(* Logix 5000 project; controller DSFW_Budzar vendor 1 type 14 code 154 rev 32.13; software revision 32.03; part 3 of 5 *)
(* tags used below, declared in another part *)
   ALARMS : DINT[5];
   ALWAYS_OFF : BOOL;
   Batch_Mode_Enable : BOOL;
   BudLib_P2T_1 : BudLib_Superheat_Subcooling;
   BudLib_P2T_2 : BudLib_Superheat_Subcooling;
   BudLib_P2T_3 : BudLib_Superheat_Subcooling;
   CLR_Alarms : BOOL;
   Compressor_R404A_Subcooling : REAL;
   Compressor_R404A_Superheat : REAL;
   CR_108 : ALIAS FOR Local:1:O.Data.0;   // Process Pump Motor Relay (Energizes Contactor M-101)
   CR_109 : ALIAS FOR Local:1:O.Data.5;   // Compressor Motor Relay (Energizes Contactor C-101)
   CR_201 : ALIAS FOR Local:1:O.Data.8;   // GFS-10 Auto Start Relay (Enables Glycol Pump)
   Enable_Batch : BOOL;   // Batch/Jacket Mode 0=Jacket 1=Batch
   Evaporator_R404A_Superheat : REAL;
   F8 : REAL[48];   // FLOAT DATA FOR PLANT SUPERVISORY SYSTEM
   FIC_101_Run_PID : BOOL;
   FIC_101_Stop_PID : BOOL;
   FIT_101 : BL_Analog_Input;   // Flow Indicating Transmitter
   FIT_101_PID_Scale_Max : REAL;
   FIT_101_PID_Scale_Min : REAL;
   Glycol_Pump_Disable_TMR : TIMER;   // Disable Glycol Fill Pump on High PSI (backup for Pressure Switch on Neptune)
   HMI_Bypass_Speed : DINT;
   HMI_Bypass_Status : BOOL;
   HMI_FCV_101_CV : REAL;
   HMI_Heater_1_Lamp : BOOL;
   HMI_Pump_Start : BOOL;
   HMI_Pump_Status : BOOL;
   HMI_Pump_Stop : BOOL;
   HMI_Ramping : BOOL;
   HMI_SCR_Max : DINT;
   HMI_Soaking : BOOL;
   HMI_Supply_Flow_Speed : DINT;
   HMI_Supply_Flow_Status : BOOL;
   Local_System_Start : BOOL;   // Local System Start 0=Stop 1=Start
   Local_Temp_Setpoint : REAL;   // Local Temperature Setpoint
   M_101_AUX : ALIAS FOR Local:1:I.Data.3;
   ONS : DINT[3];   // One-Shots
   PLC_DateTime : DINT[7];
   PM_101 : ALIAS FOR Local:1:I.Data.1;
   PT_101 : BL_Analog_Input;   // Process Supply Pressure
   PT_102 : BL_Analog_Input;   // R404A Compressor Suction Pressure
   PT_102_PID_Scale_Max : REAL;
   PT_102_PID_Scale_Min : REAL;
   PT_103 : BL_Analog_Input;   // R404A Compressor Discharge Pressure
   PT_103_PID_Scale_Max : REAL;
   PT_103_PID_Scale_Min : REAL;
   PT_104 : BL_Analog_Input;   // R404A Evaporator Suction Pressure
   PT_104_PID_Scale_Max : REAL;
   PT_104_PID_Scale_Min : REAL;
   PT_105 : BL_Analog_Input;   // Condenser Chilled Glycol Return Pressure
   PT_106 : BL_Analog_Input;   // Condenser Chilled Glycol Supply Pressure
   PT_107 : BL_Analog_Input;   // Process Pump Suction Pressure
   PT_108 : BL_Analog_Input;   // Process Pump Suction Discharge Pressure
   Pump_Manual_Release : BOOL;
   Pump_Manual_Release_Timer : TIMER;
   Pump_OK_To_Run : BOOL;
   REACTOR_BATCH_PID_START : BOOL;
   REACTOR_BATCH_PID_STOP : BOOL;
   REACTOR_BATCH_PIDE : PID_ENHANCED;
   REACTOR_BATCH_PV : REAL;
   REACTOR_BATCH_SP_HIGH : REAL;
   REACTOR_BATCH_SP_LOW : REAL;
   REACTOR_HEAT_RUN_PIDE : BOOL;
   REACTOR_HEAT_STOP_PIDE : BOOL;
   REACTOR_HEATERS_OK_TO_RUN : BOOL;
   REACTOR_HEATERS_TEMPERATURE_PIDE : PID_ENHANCED;
   Remote_Enable_Batch : BOOL;   // Remote Jacket/Batch Control (0=Jacket, 1=Batch)
   Remote_System_Start : BOOL;   // Remote Start/Stop 0=Stop 1=Start
   Remote_Temp_Setpoint : REAL;   // Remote Temperature Setpoint
   RX_Profile_Stop_SP_Control : TIMER;
   RX_RMPS : RAMP_SOAK;
   RX_RMPS_Current_Segment : DINT;
   RX_RMPS_Output : REAL;
   RX_RMPS_Soak_Time : REAL[11];
   RX_RMPS_Soak_Value : REAL[11];
   RX_RMPS_SP_Out : REAL;
   RX_Run_Temp_Profile : BOOL;
   RX_Start_Temperature_Profile : BOOL;
   RX_Stop_Temp_Profile : BOOL;
   SCR_Output_Percent : DINT;
   SCR_PID_Request : REAL;
   Sensor_1 : BudLib_Analog_Sensor;
   Sensor_2 : BudLib_Analog_Sensor;
   Sensor_3 : BudLib_Analog_Sensor;
   Sensor_4 : BudLib_Analog_Sensor;
   Sensor_5 : BudLib_Analog_Sensor;
   Sensor_6 : BudLib_Analog_Sensor;
   Sensor_7 : BudLib_Analog_Sensor;
   Sensor_8 : BudLib_Analog_Sensor;
   Sensor_9 : BudLib_Analog_Sensor;
   System_Mode : BOOL;   // 0 = Local Control 1 = Remote Control
   System_Start : BOOL;   // System Start
   T_SENSOR_1 : BudLib_Analog_Sensor;
   T_SENSOR_2 : BudLib_Analog_Sensor;
   T_SENSOR_3 : BudLib_Analog_Sensor;
   T_SENSOR_4 : BudLib_Analog_Sensor;
   T_SENSOR_5 : BudLib_Analog_Sensor;
   T_SENSOR_6 : BudLib_Analog_Sensor;
   T_SENSOR_8 : BudLib_Analog_Sensor;
   TE_101 : BL_Analog_Input;   // Process Supply Temperature
   TE_102 : BL_Analog_Input;   // Process Return Temperature
   TE_103 : BL_Analog_Input;   // R507A Liquid Line Temperature
   TE_104 : BL_Analog_Input;   // R507A Evaporator Suction Temperature
   TE_105 : BL_Analog_Input;   // R507A Compressor Suction Temperature
   TE_106 : BL_Analog_Input;   // CONDENSER CHILLED GLYCOL OUTLET TEMPERATURE SENSOR
   TE_108 : BL_Analog_Input;   // CONDENSER CHILLED GLYCOL INLET TEMPERATURE SENSOR
   Temperature_Setpoint : REAL;
   Temperature_Setpoint_Max : REAL;   // Maximum Operating Temperature Setpoint (Deg C)
   Temperature_Setpoint_Min : REAL;   // Minimum Operating Temperature Setpoint (Deg C)
   TSH_101 : ALIAS FOR Local:1:I.Data.4;
   VESSEL_TEMPERATURE : BL_Analog_Input;   // End User Reactor Temperature
(* A_MainProgram, continued *)

ROUTINE Routine_Schedule   (* ladder *)
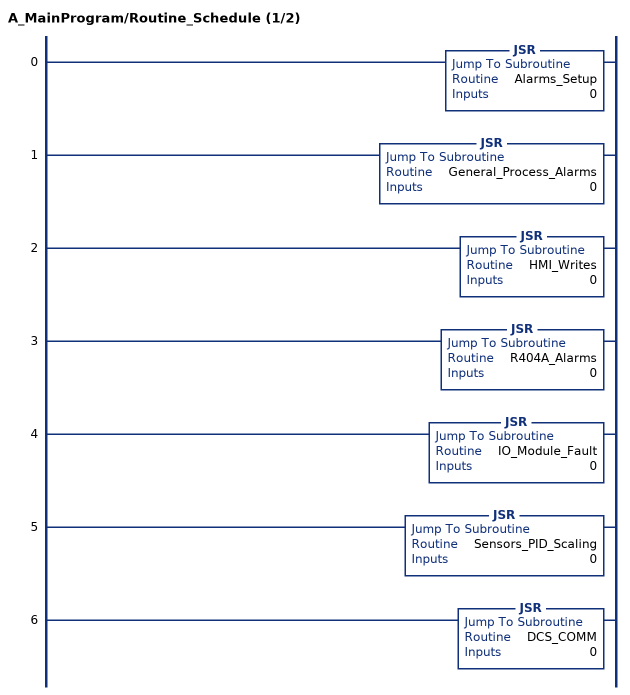
   0: JSR(Alarms_Setup,0);
   1: JSR(General_Process_Alarms,0);
   2: JSR(HMI_Writes,0);
   3: JSR(R404A_Alarms,0);
   4: JSR(IO_Module_Fault,0);
   5: JSR(Sensors_PID_Scaling,0);
   6: JSR(DCS_COMM,0);
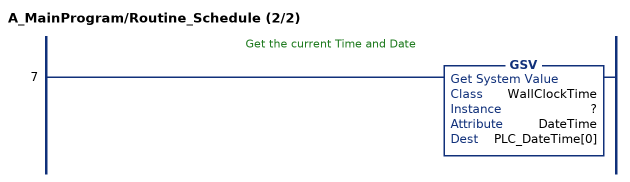
   // Get the current Time and Date
   7: GSV(WallClockTime,?,DateTime,PLC_DateTime[0]);
END_ROUTINE

ROUTINE Sensors_PID_Scaling   (* ladder *)
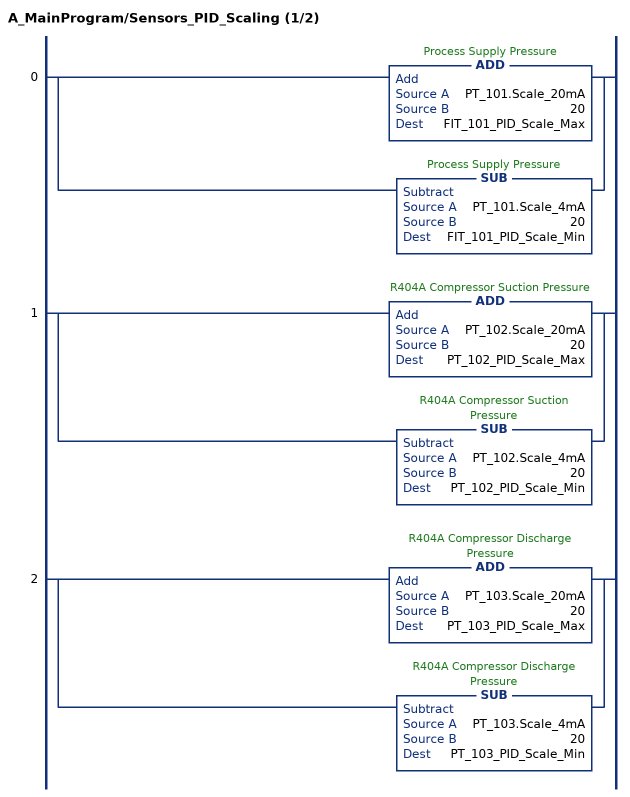
   0: [ADD(PT_101.Scale_20mA,20,FIT_101_PID_Scale_Max) ,SUB(PT_101.Scale_4mA,20,FIT_101_PID_Scale_Min) ];
   1: [ADD(PT_102.Scale_20mA,20,PT_102_PID_Scale_Max) ,SUB(PT_102.Scale_4mA,20,PT_102_PID_Scale_Min) ];
   2: [ADD(PT_103.Scale_20mA,20,PT_103_PID_Scale_Max) ,SUB(PT_103.Scale_4mA,20,PT_103_PID_Scale_Min) ];
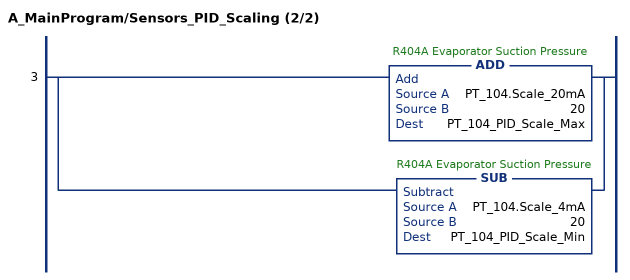
   3: [ADD(PT_104.Scale_20mA,20,PT_104_PID_Scale_Max) ,SUB(PT_104.Scale_4mA,20,PT_104_PID_Scale_Min) ];
END_ROUTINE
END_PROGRAM

PROGRAM B_Process_Control   (* main routine Main *)
VAR
   test_th : BOOL;
END_VAR

ROUTINE A_Sensors   (* ladder *)
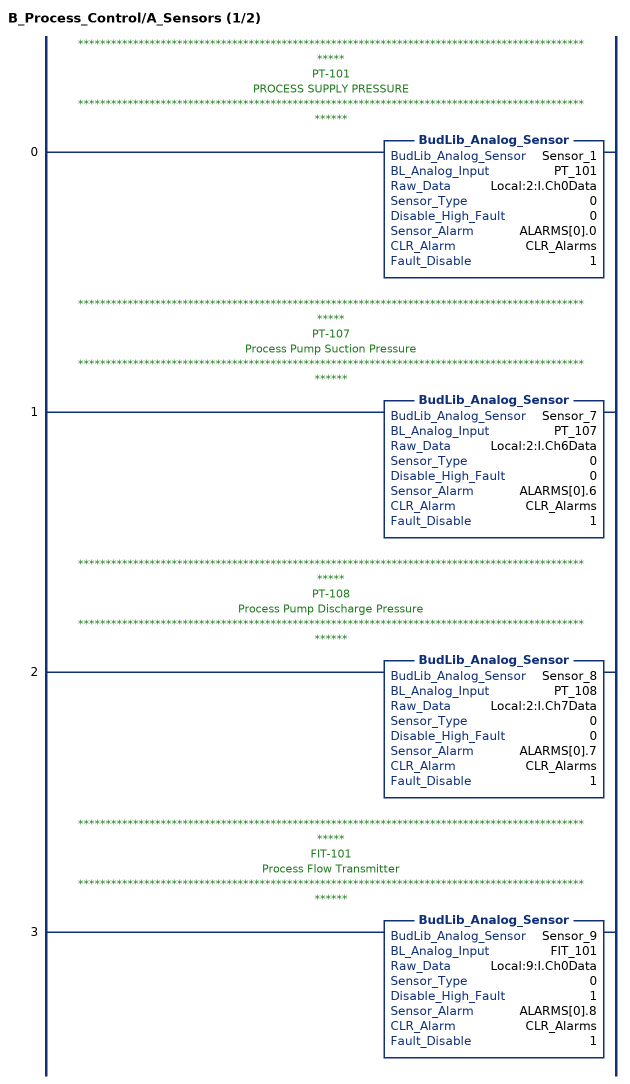
   // *************************************************************************************************
   // PT-101
   // PROCESS SUPPLY PRESSURE
   // **************************************************************************************************
   0: BudLib_Analog_Sensor(Sensor_1,PT_101,Local:2:I.Ch0Data,0,0,ALARMS[0].0,CLR_Alarms,1);
   // *************************************************************************************************
   // PT-107
   // Process Pump Suction Pressure
   // **************************************************************************************************
   1: BudLib_Analog_Sensor(Sensor_7,PT_107,Local:2:I.Ch6Data,0,0,ALARMS[0].6,CLR_Alarms,1);
   // *************************************************************************************************
   // PT-108
   // Process Pump Discharge Pressure
   // **************************************************************************************************
   2: BudLib_Analog_Sensor(Sensor_8,PT_108,Local:2:I.Ch7Data,0,0,ALARMS[0].7,CLR_Alarms,1);
   // *************************************************************************************************
   // FIT-101
   // Process Flow Transmitter
   // **************************************************************************************************
   3: BudLib_Analog_Sensor(Sensor_9,FIT_101,Local:9:I.Ch0Data,0,1,ALARMS[0].8,CLR_Alarms,1);
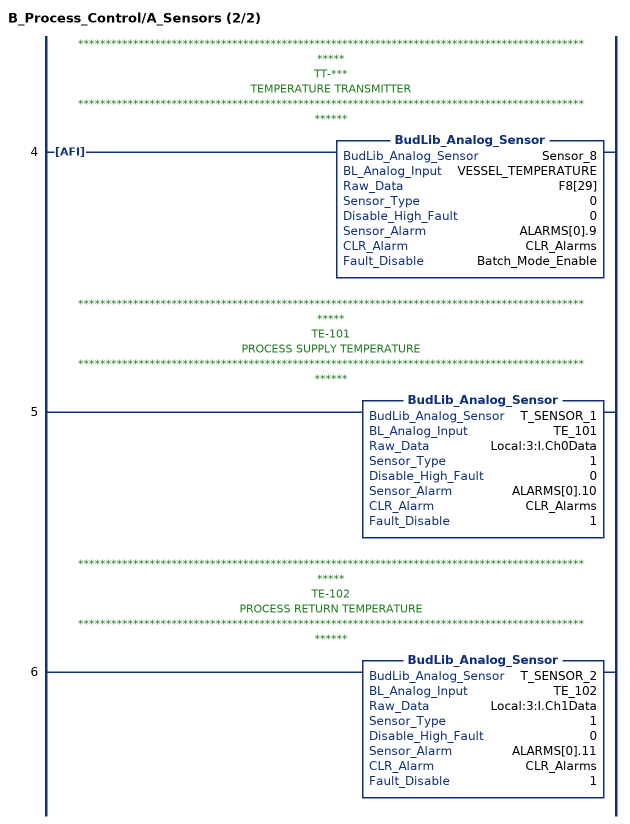
   // *************************************************************************************************
   // TT-***
   // TEMPERATURE TRANSMITTER
   // **************************************************************************************************
   4: AFI()BudLib_Analog_Sensor(Sensor_8,VESSEL_TEMPERATURE,F8[29],0,0,ALARMS[0].9,CLR_Alarms,Batch_Mode_Enable);
   // *************************************************************************************************
   // TE-101
   // PROCESS SUPPLY TEMPERATURE
   // **************************************************************************************************
   5: BudLib_Analog_Sensor(T_SENSOR_1,TE_101,Local:3:I.Ch0Data,1,0,ALARMS[0].10,CLR_Alarms,1);
   // *************************************************************************************************
   // TE-102
   // PROCESS RETURN TEMPERATURE
   // **************************************************************************************************
   6: BudLib_Analog_Sensor(T_SENSOR_2,TE_102,Local:3:I.Ch1Data,1,0,ALARMS[0].11,CLR_Alarms,1);
END_ROUTINE

ROUTINE Glycol_Tank   (* ladder *)
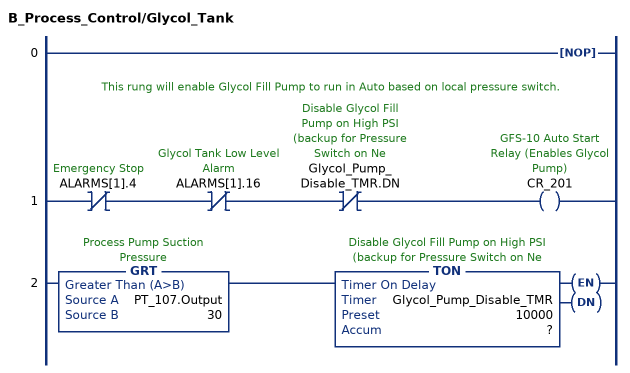
   0: NOP();
   // This rung will enable Glycol Fill Pump to run in Auto based on local pressure switch.
   1: XIO(ALARMS[1].4)XIO(ALARMS[1].16)XIO(Glycol_Pump_Disable_TMR.DN)OTE(CR_201);
   2: GRT(PT_107.Output,30)TON(Glycol_Pump_Disable_TMR,?,?);
END_ROUTINE

ROUTINE Heaters_Control   (* ladder *)
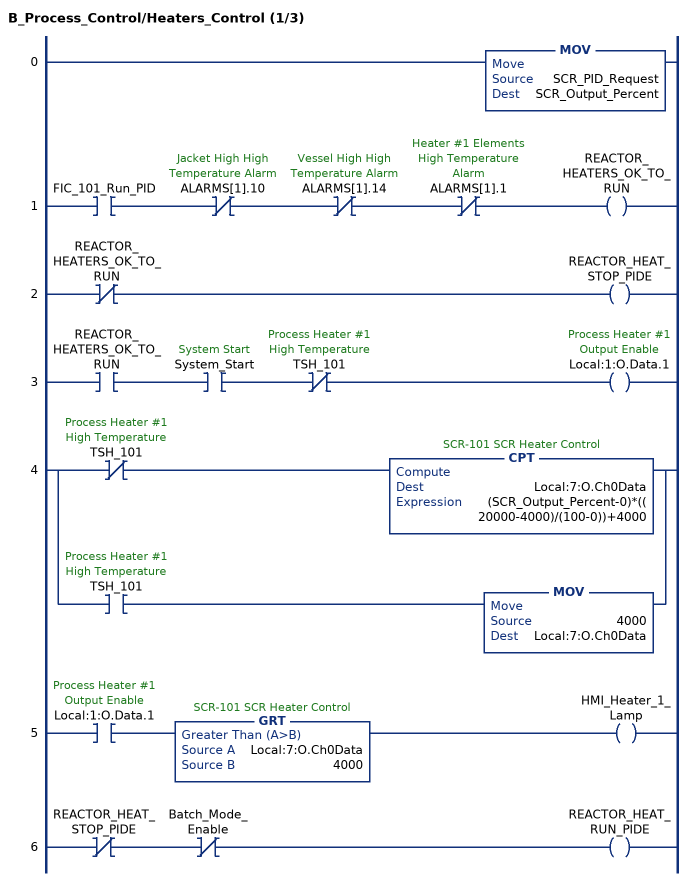
   0: MOV(SCR_PID_Request,SCR_Output_Percent);
   1: XIC(FIC_101_Run_PID)XIO(ALARMS[1].10)XIO(ALARMS[1].14)XIO(ALARMS[1].1)OTE(REACTOR_HEATERS_OK_TO_RUN);
   2: XIO(REACTOR_HEATERS_OK_TO_RUN)OTE(REACTOR_HEAT_STOP_PIDE);
   3: XIC(REACTOR_HEATERS_OK_TO_RUN)XIC(System_Start)XIO(TSH_101)OTE(Local:1:O.Data.1);
   4: [XIO(TSH_101) CPT(Local:7:O.Ch0Data,(SCR_Output_Percent-0)*((20000-4000)/(100-0))+4000) ,XIC(TSH_101) MOV(4000,Local:7:O.Ch0Data) ];
   5: XIC(Local:1:O.Data.1)GRT(Local:7:O.Ch0Data,4000)OTE(HMI_Heater_1_Lamp);
   6: XIO(REACTOR_HEAT_STOP_PIDE)XIO(Batch_Mode_Enable)OTE(REACTOR_HEAT_RUN_PIDE);
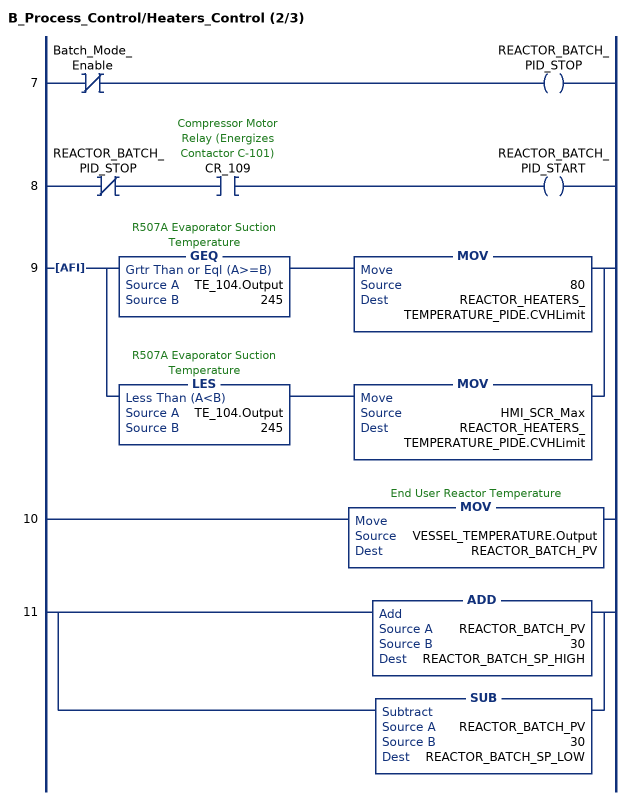
   7: XIO(Batch_Mode_Enable)OTE(REACTOR_BATCH_PID_STOP);
   8: XIO(REACTOR_BATCH_PID_STOP)XIC(CR_109)OTE(REACTOR_BATCH_PID_START);
   9: AFI()[GEQ(TE_104.Output,245) MOV(80,REACTOR_HEATERS_TEMPERATURE_PIDE.CVHLimit) ,LES(TE_104.Output,245) MOV(HMI_SCR_Max,REACTOR_HEATERS_TEMPERATURE_PIDE.CVHLimit) ];
   10: MOV(VESSEL_TEMPERATURE.Output,REACTOR_BATCH_PV);
   11: [ADD(REACTOR_BATCH_PV,30,REACTOR_BATCH_SP_HIGH) ,SUB(REACTOR_BATCH_PV,30,REACTOR_BATCH_SP_LOW) ];
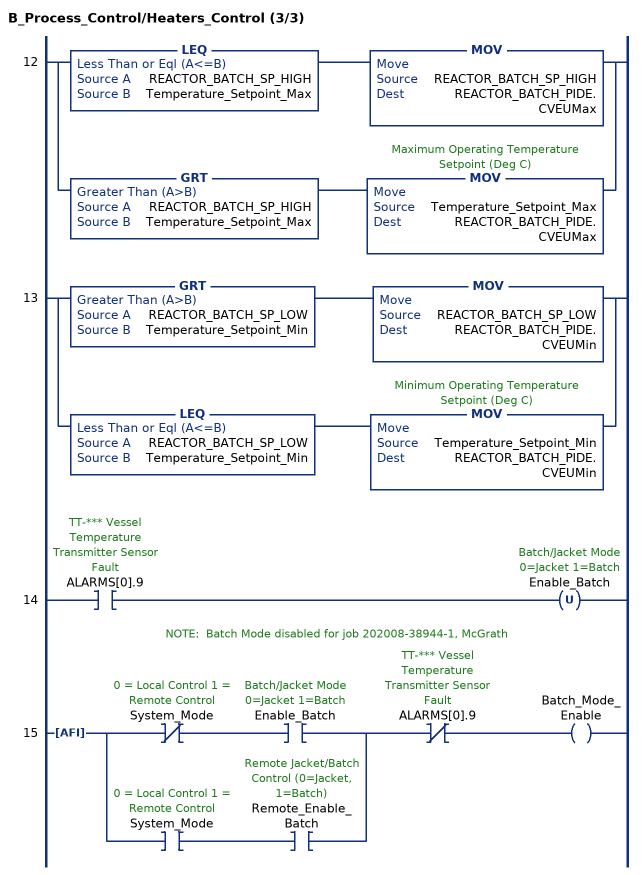
   12: [LEQ(REACTOR_BATCH_SP_HIGH,Temperature_Setpoint_Max) MOV(REACTOR_BATCH_SP_HIGH,REACTOR_BATCH_PIDE.CVEUMax) ,GRT(REACTOR_BATCH_SP_HIGH,Temperature_Setpoint_Max) MOV(Temperature_Setpoint_Max,REACTOR_BATCH_PIDE.CVEUMax) ];
   13: [GRT(REACTOR_BATCH_SP_LOW,Temperature_Setpoint_Min) MOV(REACTOR_BATCH_SP_LOW,REACTOR_BATCH_PIDE.CVEUMin) ,LEQ(REACTOR_BATCH_SP_LOW,Temperature_Setpoint_Min) MOV(Temperature_Setpoint_Min,REACTOR_BATCH_PIDE.CVEUMin) ];
   14: XIC(ALARMS[0].9)OTU(Enable_Batch);
   // NOTE:  Batch Mode disabled for job 202008-38944-1, McGrath
   15: AFI()[XIO(System_Mode) XIC(Enable_Batch) ,XIC(System_Mode) XIC(Remote_Enable_Batch) ]XIO(ALARMS[0].9)OTE(Batch_Mode_Enable);
END_ROUTINE

ROUTINE Main   (* ladder *)
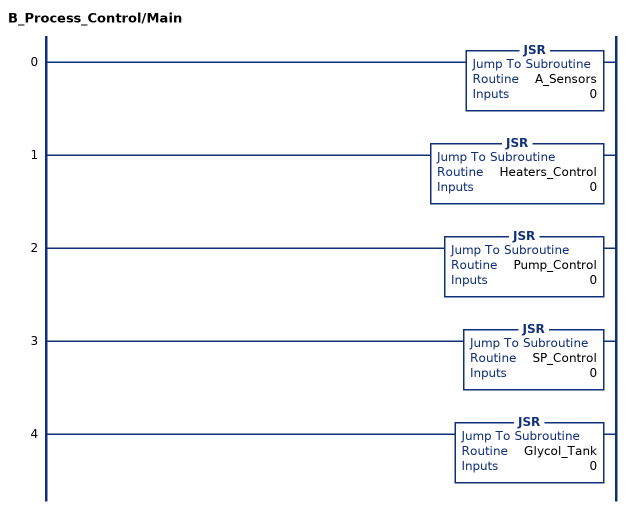
   0: JSR(A_Sensors,0);
   1: JSR(Heaters_Control,0);
   2: JSR(Pump_Control,0);
   3: JSR(SP_Control,0);
   4: JSR(Glycol_Tank,0);
END_ROUTINE

ROUTINE Pump_Control   (* ladder *)
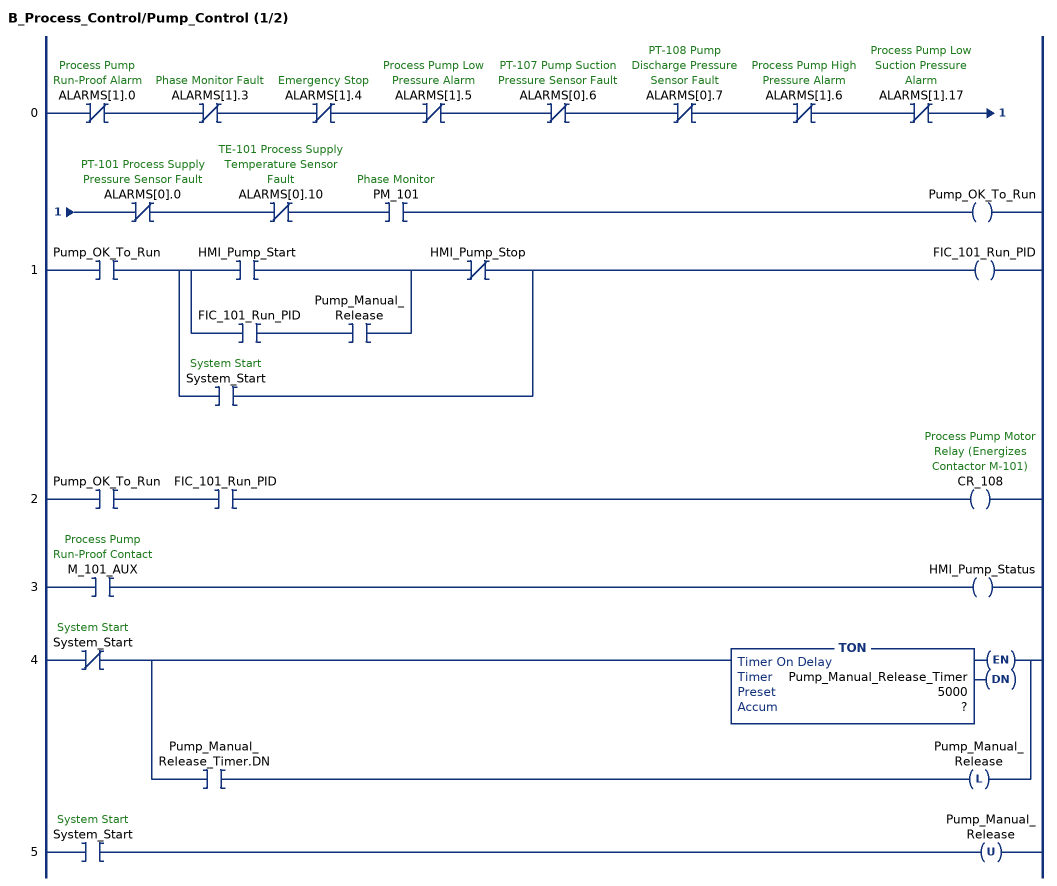
   0: XIO(ALARMS[1].0)XIO(ALARMS[1].3)XIO(ALARMS[1].4)XIO(ALARMS[1].5)XIO(ALARMS[0].6)XIO(ALARMS[0].7)XIO(ALARMS[1].6)XIO(ALARMS[1].17)XIO(ALARMS[0].0)XIO(ALARMS[0].10)XIC(PM_101)OTE(Pump_OK_To_Run);
   1: XIC(Pump_OK_To_Run)[[XIC(HMI_Pump_Start) ,XIC(FIC_101_Run_PID) XIC(Pump_Manual_Release) ] XIO(HMI_Pump_Stop) ,XIC(System_Start) ]OTE(FIC_101_Run_PID);
   2: XIC(Pump_OK_To_Run)XIC(FIC_101_Run_PID)OTE(CR_108);
   3: XIC(M_101_AUX)OTE(HMI_Pump_Status);
   4: XIO(System_Start)[TON(Pump_Manual_Release_Timer,?,?) ,XIC(Pump_Manual_Release_Timer.DN) OTL(Pump_Manual_Release) ];
   5: XIC(System_Start)OTU(Pump_Manual_Release);
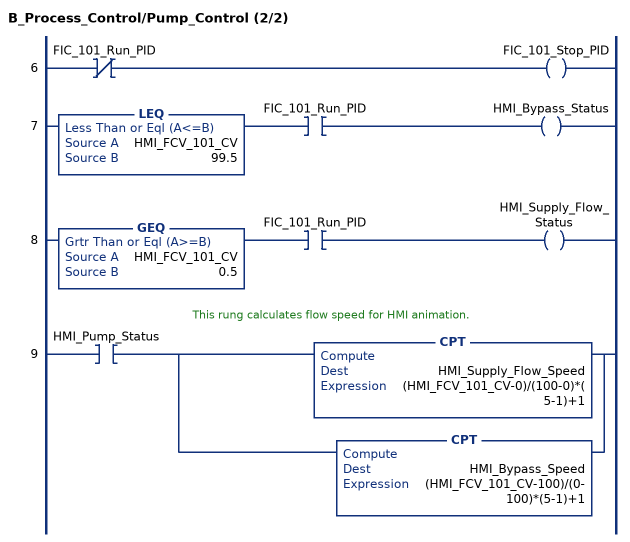
   6: XIO(FIC_101_Run_PID)OTE(FIC_101_Stop_PID);
   7: LEQ(HMI_FCV_101_CV,99.5)XIC(FIC_101_Run_PID)OTE(HMI_Bypass_Status);
   8: GEQ(HMI_FCV_101_CV,0.5)XIC(FIC_101_Run_PID)OTE(HMI_Supply_Flow_Status);
   // This rung calculates flow speed for HMI animation.
   9: XIC(HMI_Pump_Status)[CPT(HMI_Supply_Flow_Speed,(HMI_FCV_101_CV-0)/(100-0)*(5-1)+1) ,CPT(HMI_Bypass_Speed,(HMI_FCV_101_CV-100)/(0-100)*(5-1)+1) ];
END_ROUTINE

ROUTINE SP_Control   (* ladder *)
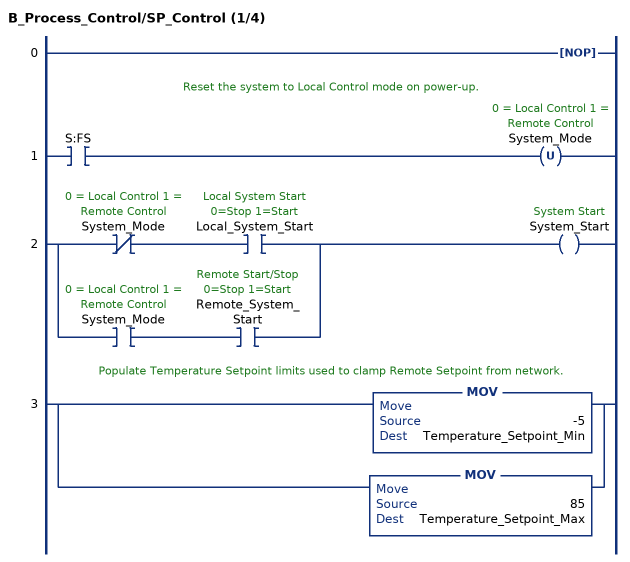
   0: NOP();
   // Reset the system to Local Control mode on power-up.
   1: XIC(S:FS)OTU(System_Mode);
   2: [XIO(System_Mode) XIC(Local_System_Start) ,XIC(System_Mode) XIC(Remote_System_Start) ]OTE(System_Start);
   // Populate Temperature Setpoint limits used to clamp Remote Setpoint from network.
   3: [MOV(-5,Temperature_Setpoint_Min) ,MOV(85,Temperature_Setpoint_Max) ];
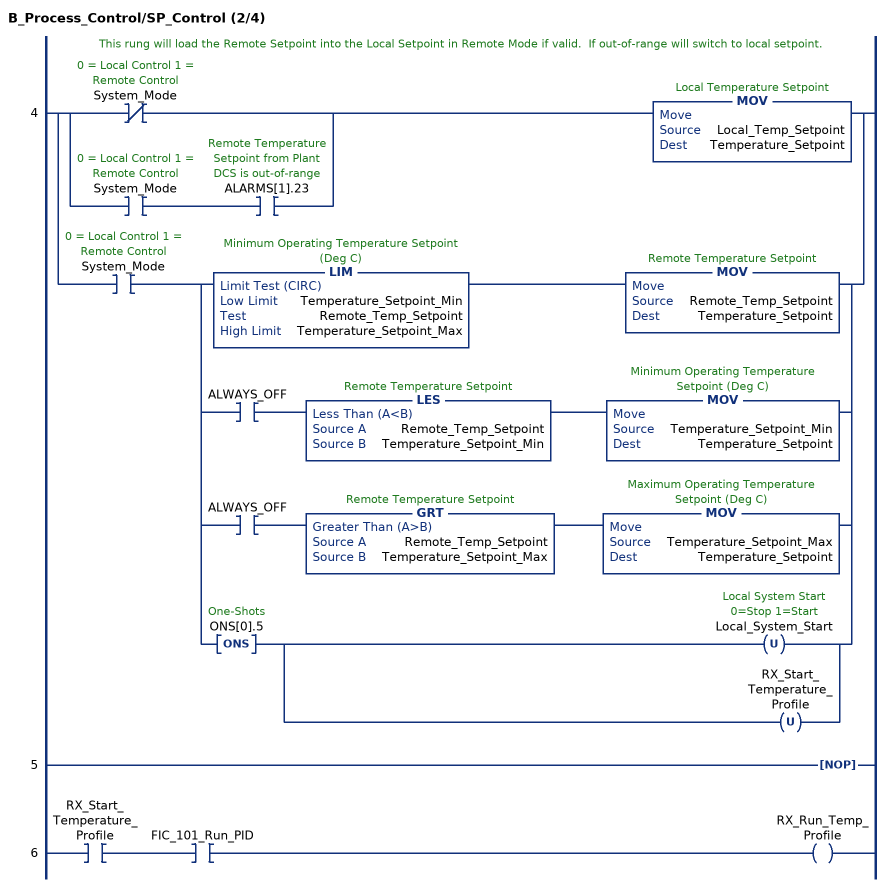
   // This rung will load the Remote Setpoint into the Local Setpoint in Remote Mode if valid.  If out-of-range will switch to local setpoint.
   4: [[XIO(System_Mode) ,XIC(System_Mode) XIC(ALARMS[1].23) ] MOV(Local_Temp_Setpoint,Temperature_Setpoint) ,XIC(System_Mode) [LIM(Temperature_Setpoint_Min,Remote_Temp_Setpoint,Temperature_Setpoint_Max) MOV(Remote_Temp_Setpoint,Temperature_Setpoint) ,XIC(ALWAYS_OFF) LES(Remote_Temp_Setpoint,Temperature_Setpoint_Min) MOV(Temperature_Setpoint_Min,Temperature_Setpoint) ,XIC(ALWAYS_OFF) GRT(Remote_Temp_Setpoint,Temperature_Setpoint_Max) MOV(Temperature_Setpoint_Max,Temperature_Setpoint) ,ONS(ONS[0].5) [OTU(Local_System_Start) ,OTU(RX_Start_Temperature_Profile) ] ] ];
   5: NOP();
   6: XIC(RX_Start_Temperature_Profile)XIC(FIC_101_Run_PID)OTE(RX_Run_Temp_Profile);
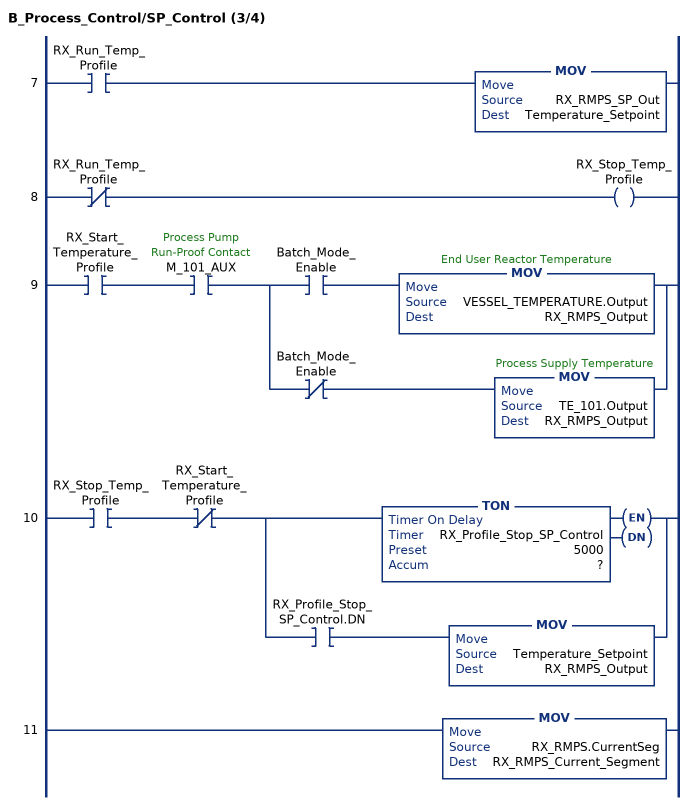
   7: XIC(RX_Run_Temp_Profile)MOV(RX_RMPS_SP_Out,Temperature_Setpoint);
   8: XIO(RX_Run_Temp_Profile)OTE(RX_Stop_Temp_Profile);
   9: XIC(RX_Start_Temperature_Profile)XIC(M_101_AUX)[XIC(Batch_Mode_Enable) MOV(VESSEL_TEMPERATURE.Output,RX_RMPS_Output) ,XIO(Batch_Mode_Enable) MOV(TE_101.Output,RX_RMPS_Output) ];
   10: XIC(RX_Stop_Temp_Profile)XIO(RX_Start_Temperature_Profile)[TON(RX_Profile_Stop_SP_Control,?,?) ,XIC(RX_Profile_Stop_SP_Control.DN) MOV(Temperature_Setpoint,RX_RMPS_Output) ];
   11: MOV(RX_RMPS.CurrentSeg,RX_RMPS_Current_Segment);
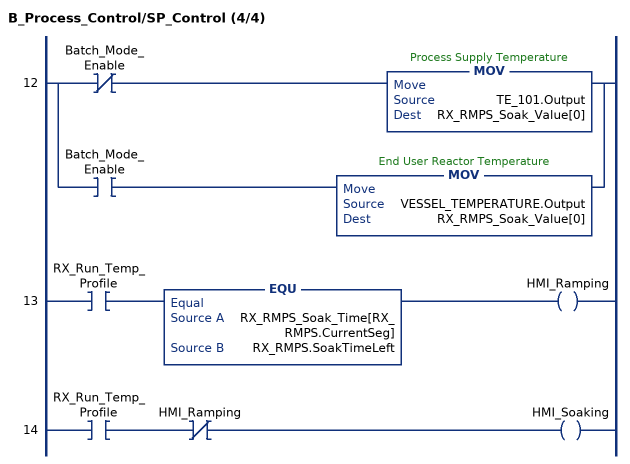
   12: [XIO(Batch_Mode_Enable) MOV(TE_101.Output,RX_RMPS_Soak_Value[0]) ,XIC(Batch_Mode_Enable) MOV(VESSEL_TEMPERATURE.Output,RX_RMPS_Soak_Value[0]) ];
   13: XIC(RX_Run_Temp_Profile)EQU(RX_RMPS_Soak_Time[RX_RMPS.CurrentSeg],RX_RMPS.SoakTimeLeft)OTE(HMI_Ramping);
   14: XIC(RX_Run_Temp_Profile)XIO(HMI_Ramping)OTE(HMI_Soaking);
END_ROUTINE
END_PROGRAM

PROGRAM D_Refrigeration_Control   (* main routine Routine_Schedule *)
VAR
   ONS1 : BOOL;
   PCV_Go_to_start_position_TMR : TIMER := (PRE := 10000, ACC := 10000);
END_VAR

ROUTINE A_Sensors   (* ladder *)
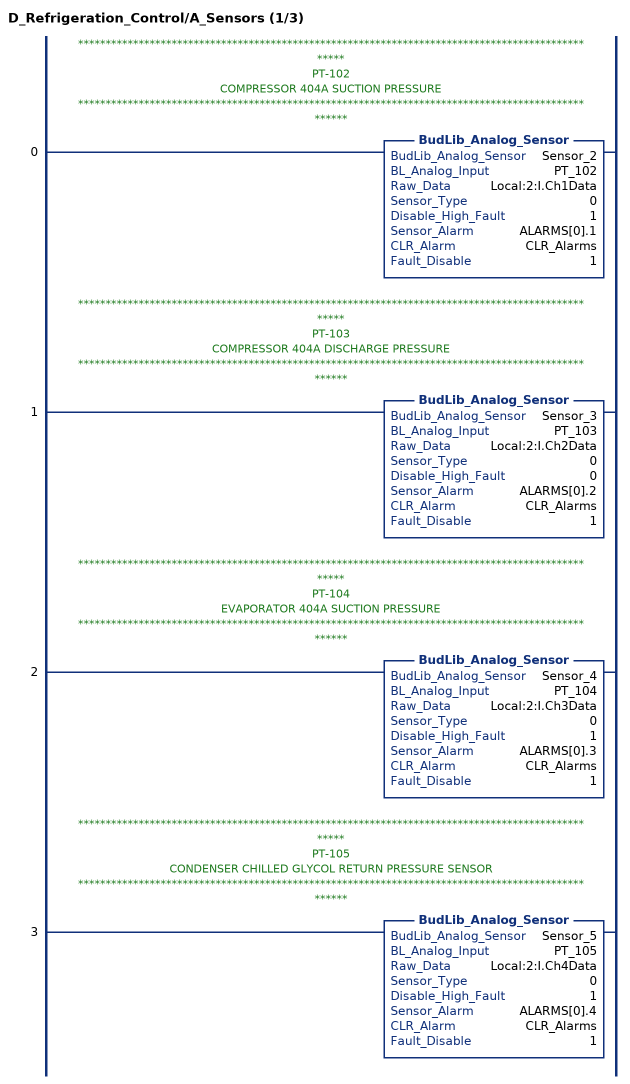
   // *************************************************************************************************
   // PT-102
   // COMPRESSOR 404A SUCTION PRESSURE
   // **************************************************************************************************
   0: BudLib_Analog_Sensor(Sensor_2,PT_102,Local:2:I.Ch1Data,0,1,ALARMS[0].1,CLR_Alarms,1);
   // *************************************************************************************************
   // PT-103
   // COMPRESSOR 404A DISCHARGE PRESSURE
   // **************************************************************************************************
   1: BudLib_Analog_Sensor(Sensor_3,PT_103,Local:2:I.Ch2Data,0,0,ALARMS[0].2,CLR_Alarms,1);
   // *************************************************************************************************
   // PT-104
   // EVAPORATOR 404A SUCTION PRESSURE
   // **************************************************************************************************
   2: BudLib_Analog_Sensor(Sensor_4,PT_104,Local:2:I.Ch3Data,0,1,ALARMS[0].3,CLR_Alarms,1);
   // *************************************************************************************************
   // PT-105
   // CONDENSER CHILLED GLYCOL RETURN PRESSURE SENSOR
   // **************************************************************************************************
   3: BudLib_Analog_Sensor(Sensor_5,PT_105,Local:2:I.Ch4Data,0,1,ALARMS[0].4,CLR_Alarms,1);
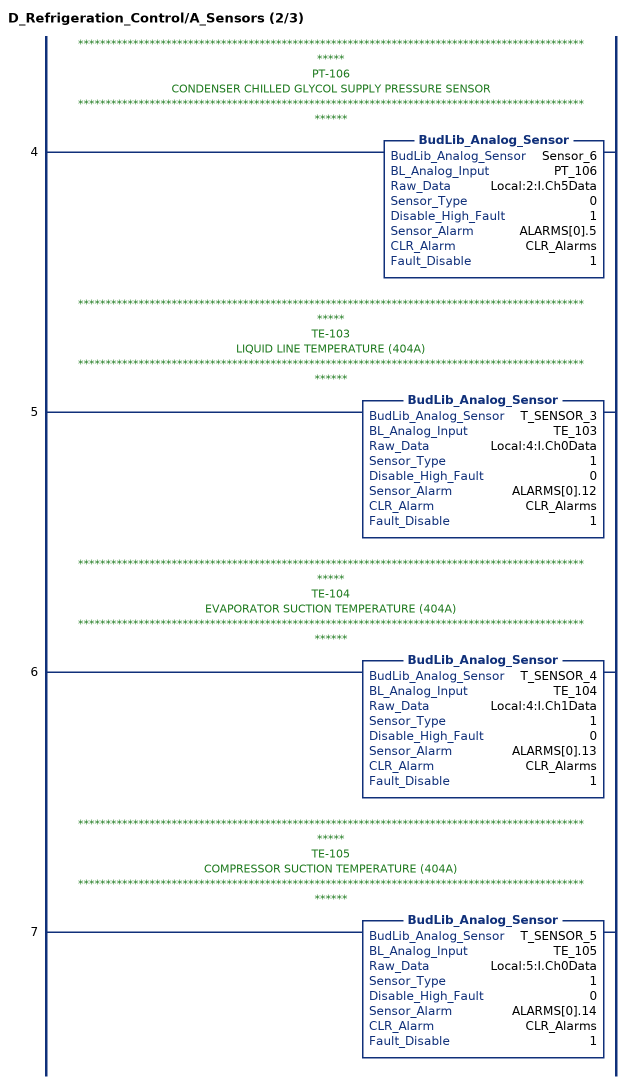
   // *************************************************************************************************
   // PT-106
   // CONDENSER CHILLED GLYCOL SUPPLY PRESSURE SENSOR
   // **************************************************************************************************
   4: BudLib_Analog_Sensor(Sensor_6,PT_106,Local:2:I.Ch5Data,0,1,ALARMS[0].5,CLR_Alarms,1);
   // *************************************************************************************************
   // TE-103
   // LIQUID LINE TEMPERATURE (404A)
   // **************************************************************************************************
   5: BudLib_Analog_Sensor(T_SENSOR_3,TE_103,Local:4:I.Ch0Data,1,0,ALARMS[0].12,CLR_Alarms,1);
   // *************************************************************************************************
   // TE-104
   // EVAPORATOR SUCTION TEMPERATURE (404A)
   // **************************************************************************************************
   6: BudLib_Analog_Sensor(T_SENSOR_4,TE_104,Local:4:I.Ch1Data,1,0,ALARMS[0].13,CLR_Alarms,1);
   // *************************************************************************************************
   // TE-105
   // COMPRESSOR SUCTION TEMPERATURE (404A)
   // **************************************************************************************************
   7: BudLib_Analog_Sensor(T_SENSOR_5,TE_105,Local:5:I.Ch0Data,1,0,ALARMS[0].14,CLR_Alarms,1);
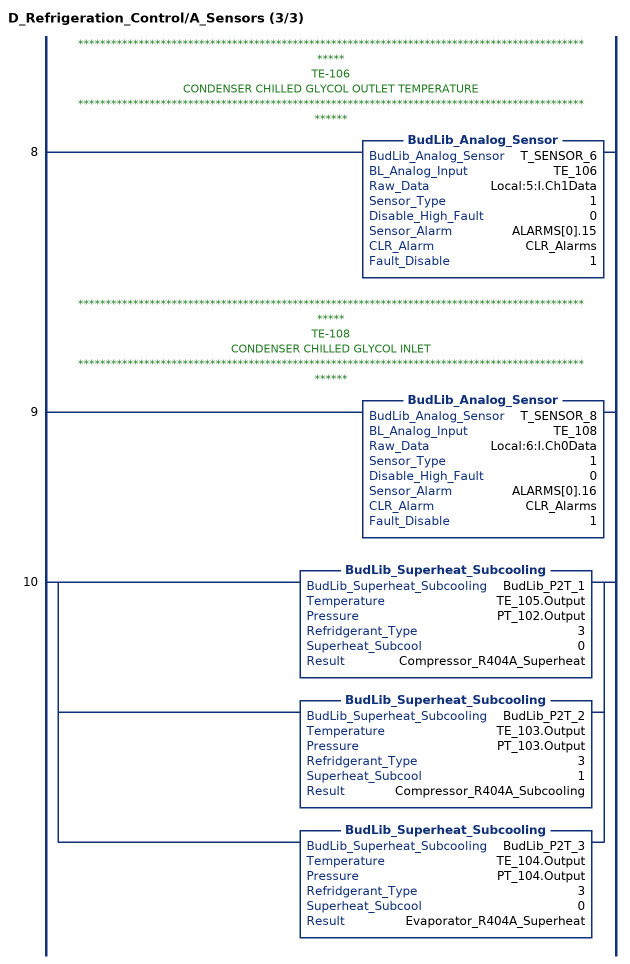
   // *************************************************************************************************
   // TE-106
   // CONDENSER CHILLED GLYCOL OUTLET TEMPERATURE
   // **************************************************************************************************
   8: BudLib_Analog_Sensor(T_SENSOR_6,TE_106,Local:5:I.Ch1Data,1,0,ALARMS[0].15,CLR_Alarms,1);
   // *************************************************************************************************
   // TE-108
   // CONDENSER CHILLED GLYCOL INLET
   // **************************************************************************************************
   9: BudLib_Analog_Sensor(T_SENSOR_8,TE_108,Local:6:I.Ch0Data,1,0,ALARMS[0].16,CLR_Alarms,1);
   10: [BudLib_Superheat_Subcooling(BudLib_P2T_1,TE_105.Output,PT_102.Output,3,0,Compressor_R404A_Superheat) ,BudLib_Superheat_Subcooling(BudLib_P2T_2,TE_103.Output,PT_103.Output,3,1,Compressor_R404A_Subcooling) ,BudLib_Superheat_Subcooling(BudLib_P2T_3,TE_104.Output,PT_104.Output,3,0,Evaporator_R404A_Superheat) ];
END_ROUTINE
